(*
SPDX-FileCopyrightText: © 2026 Oleksandr Tiutyk <trofimich@gmail.com>
SPDX-License-Identifier: MIT
License: https://opensource.org/license/mit
*)

(*!
<summary>
Beckhoff EL5002: 2-channel SSI absolute encoder interface terminal.
</summary>
<description>
Process image mapping structure for the EL5002 2-channel synchronous serial interface (SSI) absolute encoder
terminal.
Select the two-byte status PDO for each channel. The one-byte status variant is unsupported.
When used for I/O, link located fields or their containing buffers to the matching selected PDOs.
The record is not a packed wire buffer; compiler padding is not part of the device specification.
Unlinked/default values do not prove valid I/O. The caller evaluates bus/channel validity before use.
Use one owner task per instance and externally synchronize other access; multi-field snapshots are not atomic.
Copies store data without creating hardware links. Keep borrowed field references valid while consumers are bound.
This passive record performs no validation, synchronization, configuration or protocol advancement.
</description>
*)
TYPE EL5002 :
STRUCT
	Ch1 : SSI_ENCODER_CHANNEL;
	Ch2 : SSI_ENCODER_CHANNEL;
END_STRUCT
END_TYPE

(* stored: Version 1.1.0.1, ProductVersion 3.1.4026.20
   DUT EL5002: Id {9159eb16-6698-4a53-8fc2-ca57486dcfd6} *)
